ADAPTER AOption (* Optionsmanagement-Adapter: INIT-Request/Confirm-Handshake mit QI (Event Input Qualifier, IEC 61499-1) *)
  (* Standard: 61499-1; Description: Copyright (c) 2026 Meisterschulen am Ostbahnhof This program and the accompanying materials are made available under the terms of the Eclipse Public License 2.0 which is available at https://www.eclipse.org/legal/epl-2.0/ SPDX-License-Identifier: EPL-2.0 *)
  (* Version 1.0, 2026-10-13, Franz Höpfinger, Meisterschulen am Ostbahnhof, initial API and implementation and/or initial documentation *)
  PACKAGE Option;
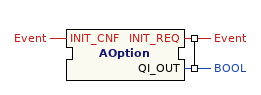
  EVENT_INPUT
    INIT_CNF; (* Initialisierung bestaetigt (SOCKET -> PLUG) *)
  END_EVENT
  EVENT_OUTPUT
    INIT_REQ WITH QI_OUT; (* Initialisierung anfordern (PLUG -> SOCKET) *)
  END_EVENT
  VAR_OUTPUT
    QI_OUT : BOOL; (* Event Input Qualifier zu INIT_REQ (IEC 61499-1): TRUE = Option anfordern/aktivieren (INIT_REQ+), FALSE = zurueckziehen/terminieren (INIT_REQ-) *)
  END_VAR
END_ADAPTER
